(* Logix 5000 project; controller CIP_14485201 vendor 1 type 14 code 216 rev 38.11; software revision 38.01; part 10 of 12 *)
(* tags used below, declared in another part *)
   Bit : BOOL[128];   // BIT
   Integer : DINT[150];   // INTEGER
   MOA_OFF : DINT[20];   // PANELVIEW MOA OFF
   MOA_ON : DINT[20];   // PANELVIEW MOA ON
   MOA_One_Shot : BOOL[32];   // PANELVIEW MOA ONE SHOT
   MOA_Screen1_Auto : BOOL;   // PV MOA SCREEN #1 AUTO PB
   MOA_Screen1_Man_Off : BOOL;   // PV MOA SCREEN #1 OFF PB
   MOA_Screen1_Man_On : BOOL;   // PV MOA SCREEN #1 MANUAL PB
   MOA_Screen2_Auto : BOOL;   // PV MOA SCREEN #2 AUTO PB
   MOA_Screen2_Man_Off : BOOL;   // PV MOA SCREEN #2 OFF PB
   MOA_Screen2_Man_On : BOOL;   // PV MOA SCREEN #2 MANUAL PB
   MOA_Select : DINT[10];   // MAN/OFF/AUTO SELECT
   MOA_Status : DINT[10];   // MAN/OFF/AUTO STATUS
   One_Shot : BOOL[128];   // ONE SHOT ARRAY
   OpCode_Pin : DINT[5];   // OPCODE PIN ARRAY
   Panelview : INT[40];   // PANELVIEW CONTROL
   Recipe : RECIPE[41];   // RECIPES
   SCLD_Return_Temp : SCALE;   // RETURN TEMPERATURE 0-100°C
   SCLD_Rinse_Cond : SCALE;   // RINSE CONDUCTIVITY 0-10 uS/cm
   SCLD_Supply_Temp : SCALE;   // SUPPLY TEMPERATURE 0-100°C
   SCLD_Wash_Cond : SCALE;   // WASH CONDUCTIVITY 0-100 mS/cm
   SP_Return_Temp : REAL;   // CURRENT RETURN TEMP SETPOINT
   SP_Rinse_Cond : REAL;   // CURRENT RINSE CONDUCTIVITY SETPOINT
   SP_Supply_Temp : REAL;   // CURRENT SUPPLY TEMP SETPOINT
   SP_Wash_Cond : REAL;   // CURRENT WASH CONDUCTIVITY SETPOINT
   SP_Wash_Cond_Hold : REAL;   // CURRENT WASH CONDUCTIVITY SETPOINT LOW HOLD
   Subsequent_OpCode_Pin : DINT[5];   // OPCODE PIN ARRAY
   Timer : TIMER[99];   // TIMER
   Timer_Chem1_Pump : TIMER[7];   // CHEM #1 CONTROL TIMERS
   Timer_Chem2_Pump : TIMER[7];   // CHEM #2 CONTROL TIMERS
(* MainProgram, continued *)

ROUTINE _30_MAN_OFF_AUTO   (* ladder *)
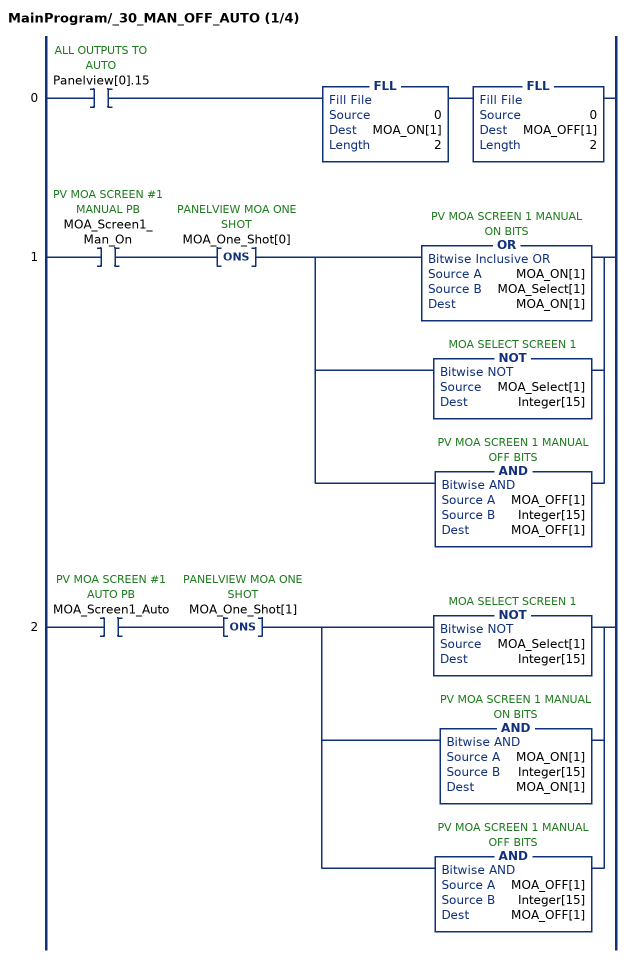
   0: XIC(Panelview[0].15)FLL(0,MOA_ON[1],2)FLL(0,MOA_OFF[1],2);
   1: XIC(MOA_Screen1_Man_On)ONS(MOA_One_Shot[0])[OR(MOA_ON[1],MOA_Select[1],MOA_ON[1]) ,NOT(MOA_Select[1],Integer[15]) ,AND(MOA_OFF[1],Integer[15],MOA_OFF[1]) ];
   2: XIC(MOA_Screen1_Auto)ONS(MOA_One_Shot[1])[NOT(MOA_Select[1],Integer[15]) ,AND(MOA_ON[1],Integer[15],MOA_ON[1]) ,AND(MOA_OFF[1],Integer[15],MOA_OFF[1]) ];
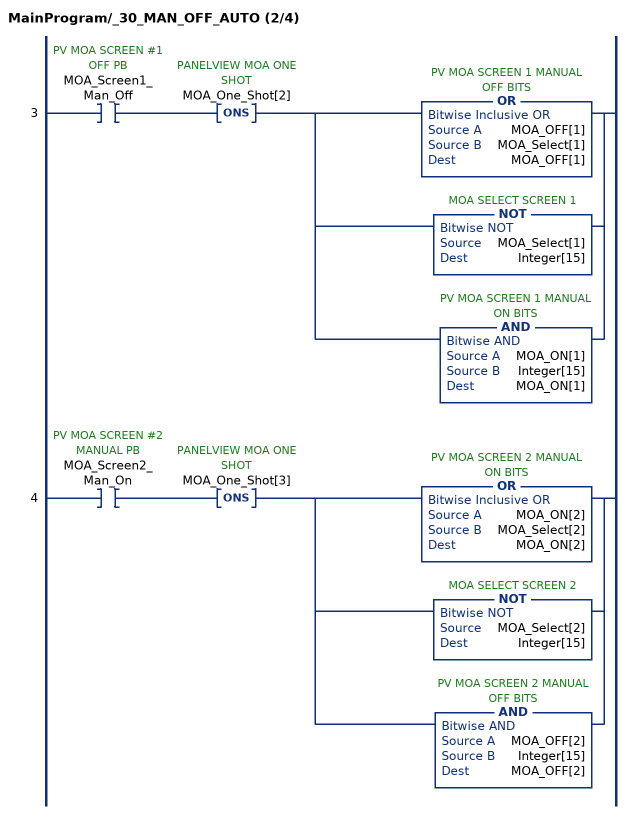
   3: XIC(MOA_Screen1_Man_Off)ONS(MOA_One_Shot[2])[OR(MOA_OFF[1],MOA_Select[1],MOA_OFF[1]) ,NOT(MOA_Select[1],Integer[15]) ,AND(MOA_ON[1],Integer[15],MOA_ON[1]) ];
   4: XIC(MOA_Screen2_Man_On)ONS(MOA_One_Shot[3])[OR(MOA_ON[2],MOA_Select[2],MOA_ON[2]) ,NOT(MOA_Select[2],Integer[15]) ,AND(MOA_OFF[2],Integer[15],MOA_OFF[2]) ];
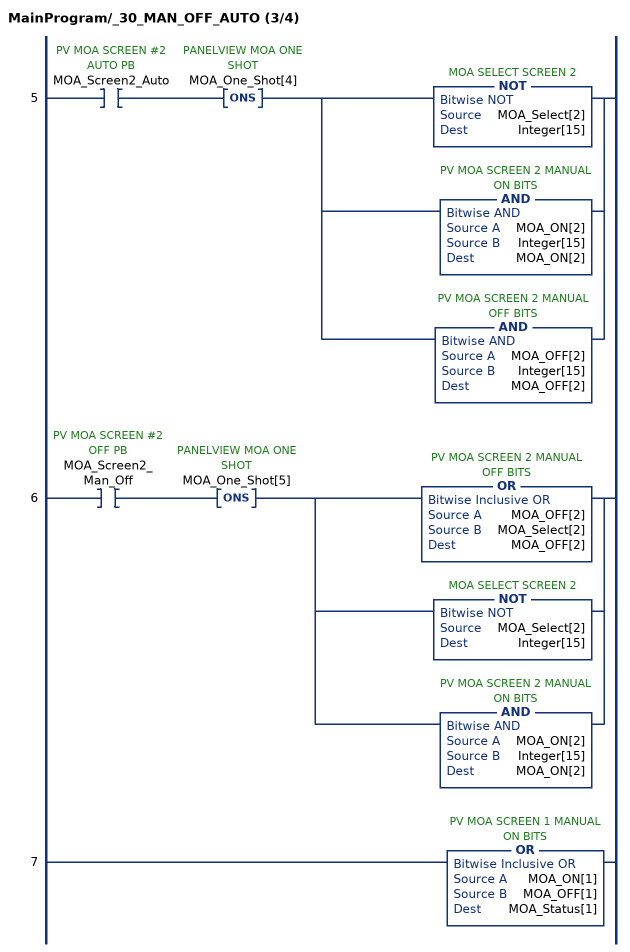
   5: XIC(MOA_Screen2_Auto)ONS(MOA_One_Shot[4])[NOT(MOA_Select[2],Integer[15]) ,AND(MOA_ON[2],Integer[15],MOA_ON[2]) ,AND(MOA_OFF[2],Integer[15],MOA_OFF[2]) ];
   6: XIC(MOA_Screen2_Man_Off)ONS(MOA_One_Shot[5])[OR(MOA_OFF[2],MOA_Select[2],MOA_OFF[2]) ,NOT(MOA_Select[2],Integer[15]) ,AND(MOA_ON[2],Integer[15],MOA_ON[2]) ];
   7: OR(MOA_ON[1],MOA_OFF[1],MOA_Status[1]);
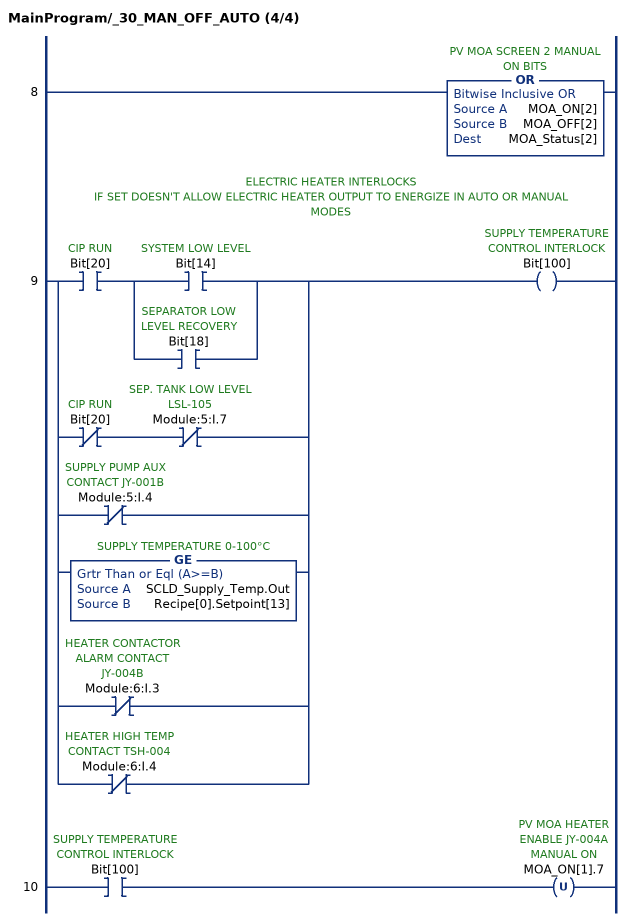
   8: OR(MOA_ON[2],MOA_OFF[2],MOA_Status[2]);
   // ELECTRIC HEATER INTERLOCKS
   // IF SET DOESN'T ALLOW ELECTRIC HEATER OUTPUT TO ENERGIZE IN AUTO OR MANUAL MODES
   9: [XIC(Bit[20]) [XIC(Bit[14]) ,XIC(Bit[18]) ] ,XIO(Bit[20]) XIO(Module:5:I.7) ,XIO(Module:5:I.4) ,GE(SCLD_Supply_Temp.Out,Recipe[0].Setpoint[13]) ,XIO(Module:6:I.3) ,XIO(Module:6:I.4) ]OTE(Bit[100]);
   10: XIC(Bit[100])OTU(MOA_ON[1].7);
END_ROUTINE

ROUTINE _86_TEMPERATURE   (* ladder *)
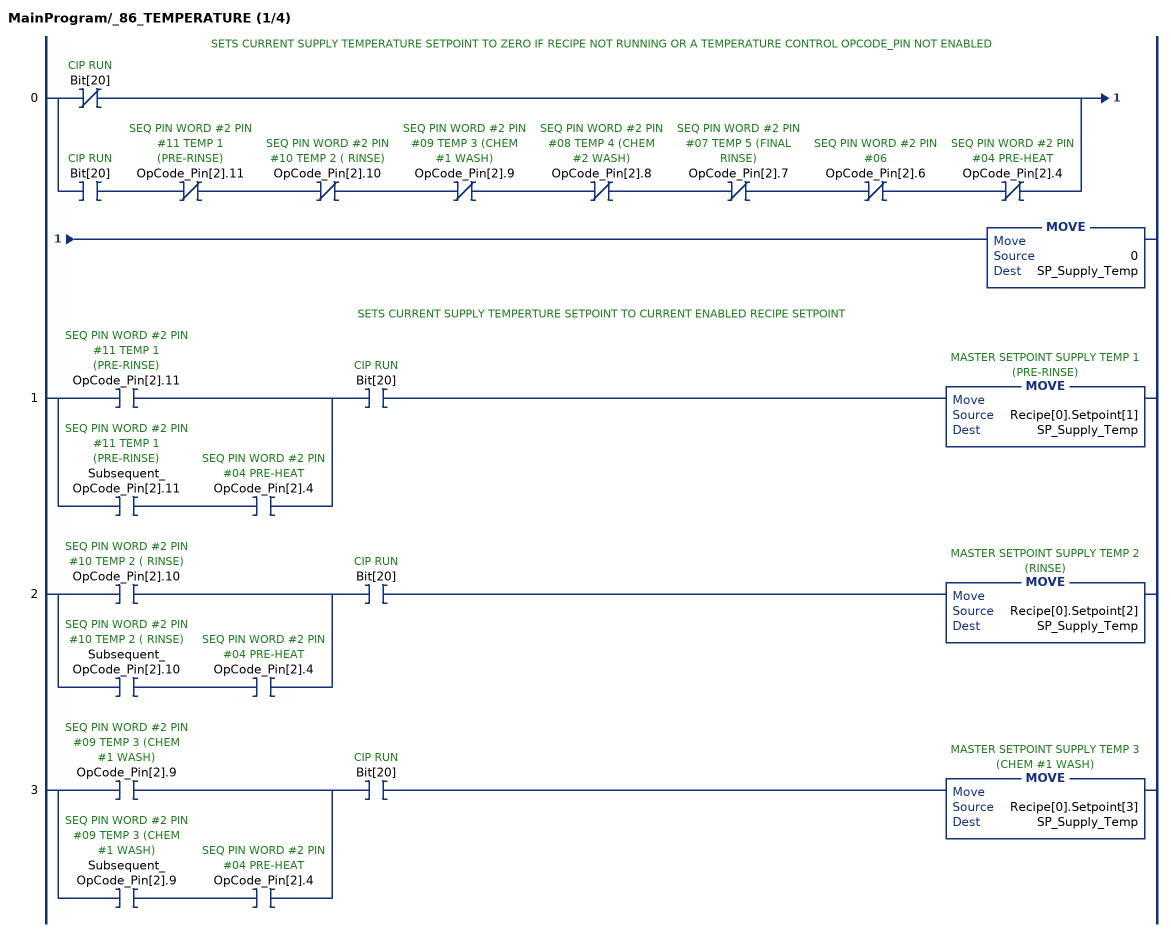
   // SETS CURRENT SUPPLY TEMPERATURE SETPOINT TO ZERO IF RECIPE NOT RUNNING OR A TEMPERATURE CONTROL OPCODE_PIN NOT ENABLED
   0: [XIO(Bit[20]) ,XIC(Bit[20]) XIO(OpCode_Pin[2].11) XIO(OpCode_Pin[2].10) XIO(OpCode_Pin[2].9) XIO(OpCode_Pin[2].8) XIO(OpCode_Pin[2].7) XIO(OpCode_Pin[2].6) XIO(OpCode_Pin[2].4) ]MOVE(0,SP_Supply_Temp);
   // SETS CURRENT SUPPLY TEMPERTURE SETPOINT TO CURRENT ENABLED RECIPE SETPOINT
   1: [XIC(OpCode_Pin[2].11) ,XIC(Subsequent_OpCode_Pin[2].11) XIC(OpCode_Pin[2].4) ]XIC(Bit[20])MOVE(Recipe[0].Setpoint[1],SP_Supply_Temp);
   2: [XIC(OpCode_Pin[2].10) ,XIC(Subsequent_OpCode_Pin[2].10) XIC(OpCode_Pin[2].4) ]XIC(Bit[20])MOVE(Recipe[0].Setpoint[2],SP_Supply_Temp);
   3: [XIC(OpCode_Pin[2].9) ,XIC(Subsequent_OpCode_Pin[2].9) XIC(OpCode_Pin[2].4) ]XIC(Bit[20])MOVE(Recipe[0].Setpoint[3],SP_Supply_Temp);
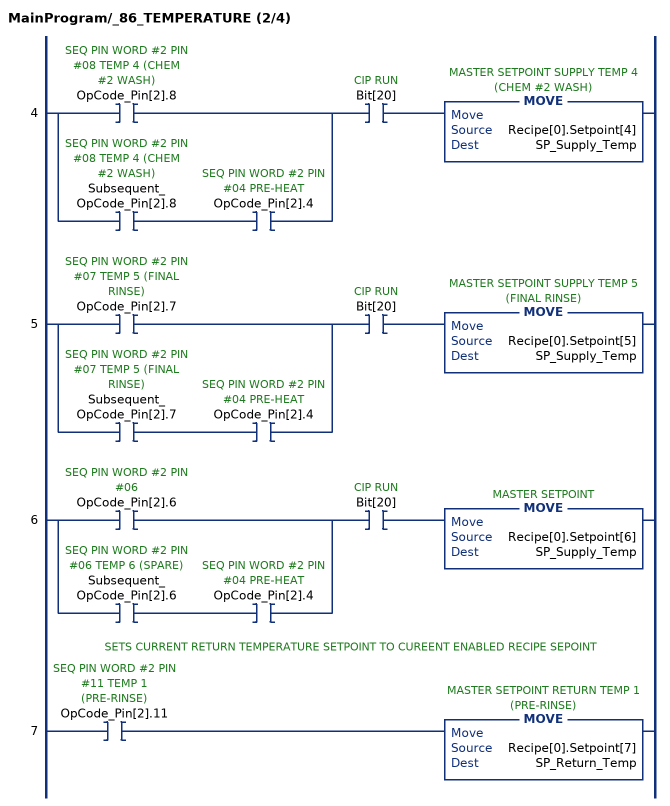
   4: [XIC(OpCode_Pin[2].8) ,XIC(Subsequent_OpCode_Pin[2].8) XIC(OpCode_Pin[2].4) ]XIC(Bit[20])MOVE(Recipe[0].Setpoint[4],SP_Supply_Temp);
   5: [XIC(OpCode_Pin[2].7) ,XIC(Subsequent_OpCode_Pin[2].7) XIC(OpCode_Pin[2].4) ]XIC(Bit[20])MOVE(Recipe[0].Setpoint[5],SP_Supply_Temp);
   6: [XIC(OpCode_Pin[2].6) ,XIC(Subsequent_OpCode_Pin[2].6) XIC(OpCode_Pin[2].4) ]XIC(Bit[20])MOVE(Recipe[0].Setpoint[6],SP_Supply_Temp);
   // SETS CURRENT RETURN TEMPERATURE SETPOINT TO CUREENT ENABLED RECIPE SEPOINT
   7: XIC(OpCode_Pin[2].11)MOVE(Recipe[0].Setpoint[7],SP_Return_Temp);
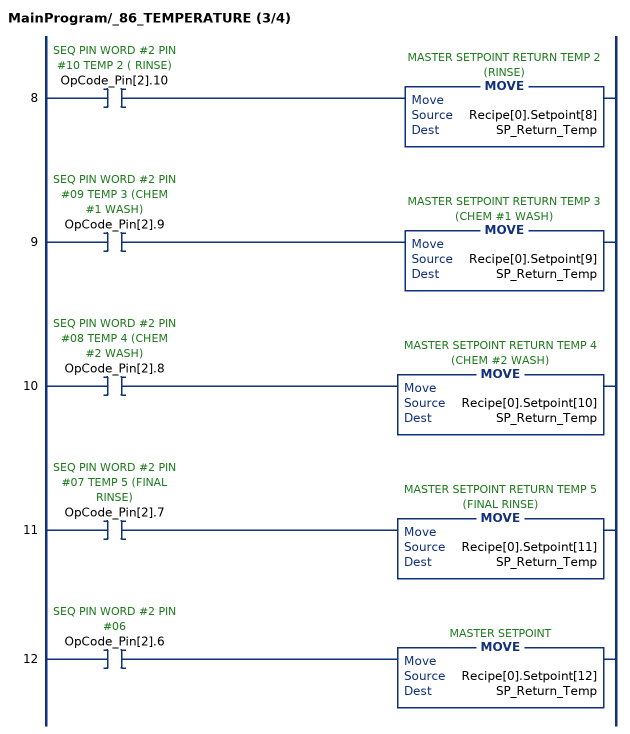
   8: XIC(OpCode_Pin[2].10)MOVE(Recipe[0].Setpoint[8],SP_Return_Temp);
   9: XIC(OpCode_Pin[2].9)MOVE(Recipe[0].Setpoint[9],SP_Return_Temp);
   10: XIC(OpCode_Pin[2].8)MOVE(Recipe[0].Setpoint[10],SP_Return_Temp);
   11: XIC(OpCode_Pin[2].7)MOVE(Recipe[0].Setpoint[11],SP_Return_Temp);
   12: XIC(OpCode_Pin[2].6)MOVE(Recipe[0].Setpoint[12],SP_Return_Temp);
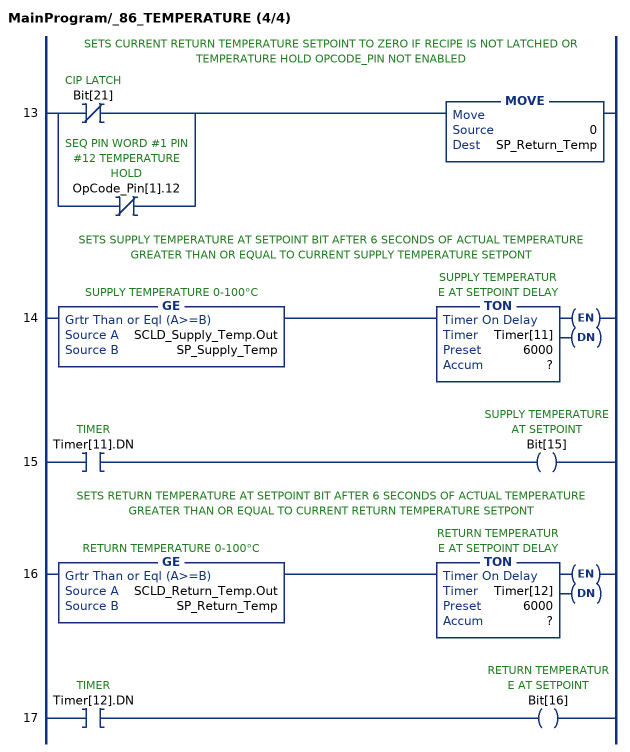
   // SETS CURRENT RETURN TEMPERATURE SETPOINT TO ZERO IF RECIPE IS NOT LATCHED OR TEMPERATURE HOLD OPCODE_PIN NOT ENABLED
   13: [XIO(Bit[21]) ,XIO(OpCode_Pin[1].12) ]MOVE(0,SP_Return_Temp);
   // SETS SUPPLY TEMPERATURE AT SETPOINT BIT AFTER 6 SECONDS OF ACTUAL TEMPERATURE GREATER THAN OR EQUAL TO CURRENT SUPPLY TEMPERATURE SETPONT
   14: GE(SCLD_Supply_Temp.Out,SP_Supply_Temp)TON(Timer[11],?,?);
   15: XIC(Timer[11].DN)OTE(Bit[15]);
   // SETS RETURN TEMPERATURE AT SETPOINT BIT AFTER 6 SECONDS OF ACTUAL TEMPERATURE GREATER THAN OR EQUAL TO CURRENT RETURN TEMPERATURE SETPONT
   16: GE(SCLD_Return_Temp.Out,SP_Return_Temp)TON(Timer[12],?,?);
   17: XIC(Timer[12].DN)OTE(Bit[16]);
END_ROUTINE

ROUTINE _87_CHEM1_PUMP   (* ladder *)
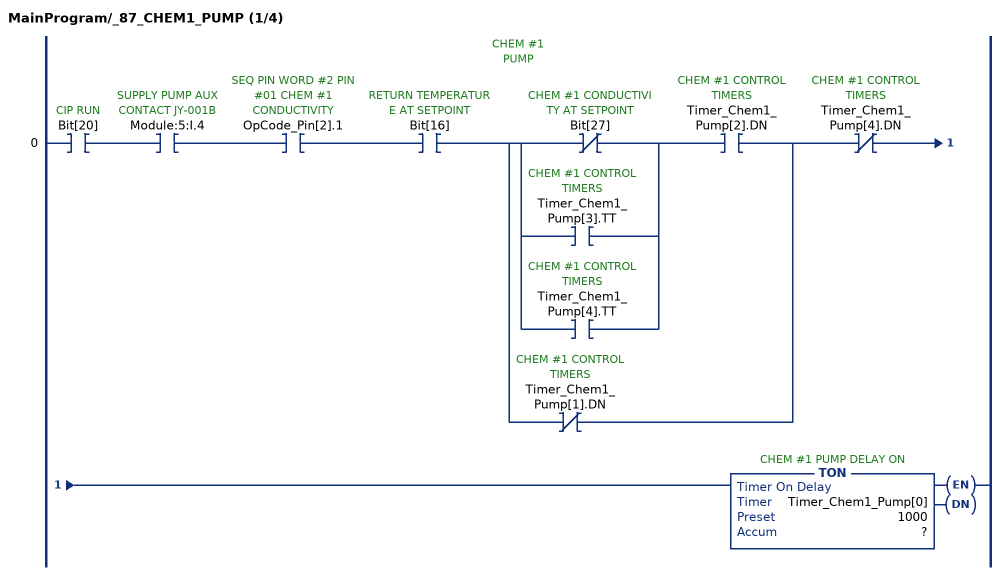
   // CHEM #1
   // PUMP
   0: XIC(Bit[20])XIC(Module:5:I.4)XIC(OpCode_Pin[2].1)XIC(Bit[16])[[XIO(Bit[27]) ,XIC(Timer_Chem1_Pump[3].TT) ,XIC(Timer_Chem1_Pump[4].TT) ] XIC(Timer_Chem1_Pump[2].DN) ,XIO(Timer_Chem1_Pump[1].DN) ]XIO(Timer_Chem1_Pump[4].DN)TON(Timer_Chem1_Pump[0],?,?);
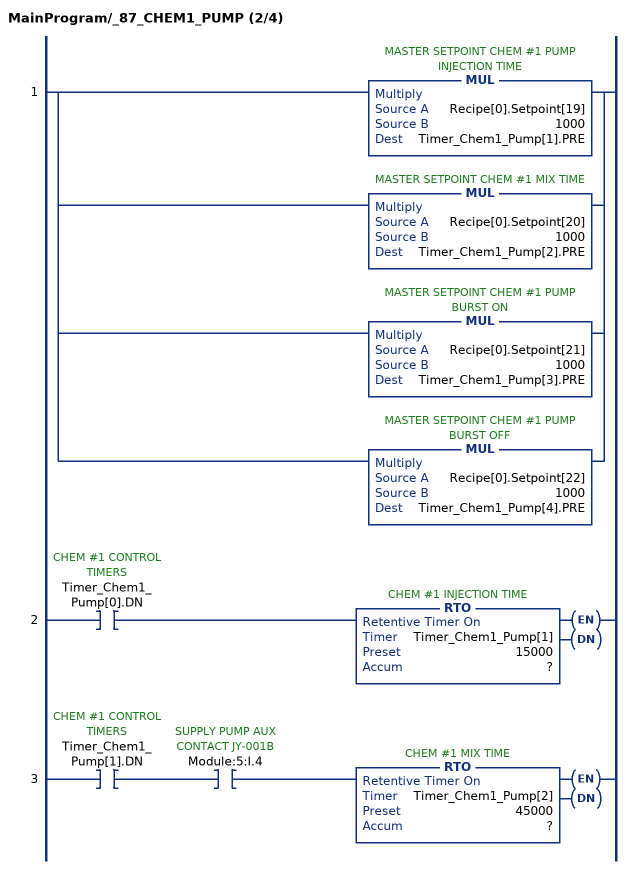
   1: [MUL(Recipe[0].Setpoint[19],1000,Timer_Chem1_Pump[1].PRE) ,MUL(Recipe[0].Setpoint[20],1000,Timer_Chem1_Pump[2].PRE) ,MUL(Recipe[0].Setpoint[21],1000,Timer_Chem1_Pump[3].PRE) ,MUL(Recipe[0].Setpoint[22],1000,Timer_Chem1_Pump[4].PRE) ];
   2: XIC(Timer_Chem1_Pump[0].DN)RTO(Timer_Chem1_Pump[1],?,?);
   3: XIC(Timer_Chem1_Pump[1].DN)XIC(Module:5:I.4)RTO(Timer_Chem1_Pump[2],?,?);
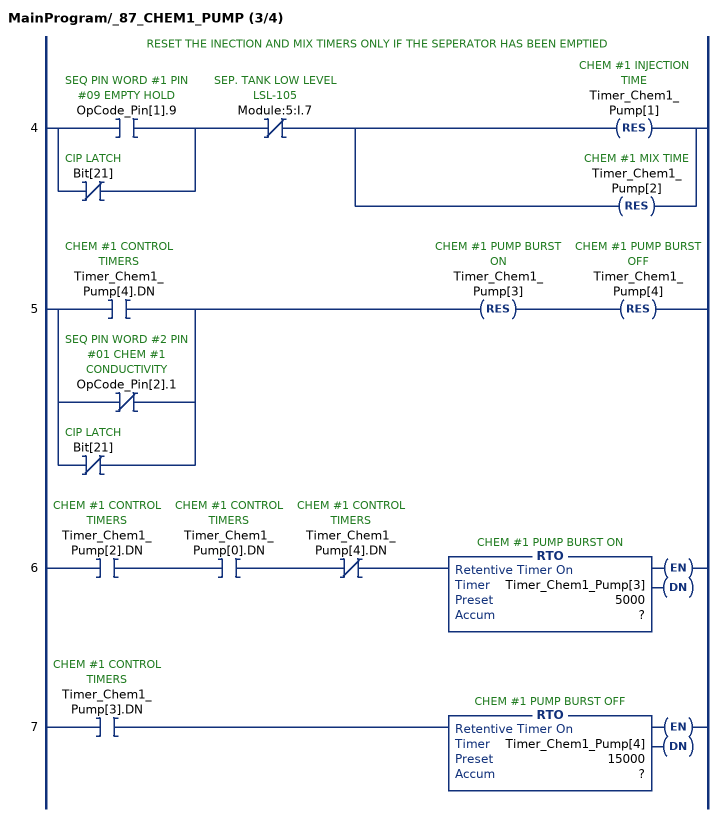
   // RESET THE INECTION AND MIX TIMERS ONLY IF THE SEPERATOR HAS BEEN EMPTIED
   4: [XIC(OpCode_Pin[1].9) ,XIO(Bit[21]) ]XIO(Module:5:I.7)[RES(Timer_Chem1_Pump[1]) ,RES(Timer_Chem1_Pump[2]) ];
   5: [XIC(Timer_Chem1_Pump[4].DN) ,XIO(OpCode_Pin[2].1) ,XIO(Bit[21]) ]RES(Timer_Chem1_Pump[3])RES(Timer_Chem1_Pump[4]);
   6: XIC(Timer_Chem1_Pump[2].DN)XIC(Timer_Chem1_Pump[0].DN)XIO(Timer_Chem1_Pump[4].DN)RTO(Timer_Chem1_Pump[3],?,?);
   7: XIC(Timer_Chem1_Pump[3].DN)RTO(Timer_Chem1_Pump[4],?,?);
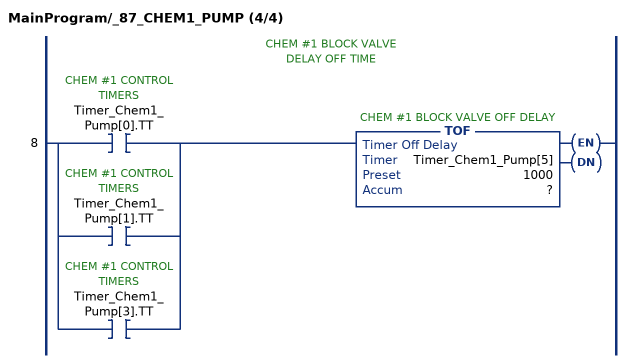
   // CHEM #1 BLOCK VALVE
   //  DELAY OFF TIME
   8: [XIC(Timer_Chem1_Pump[0].TT) ,XIC(Timer_Chem1_Pump[1].TT) ,XIC(Timer_Chem1_Pump[3].TT) ]TOF(Timer_Chem1_Pump[5],?,?);
END_ROUTINE

ROUTINE _87_CHEM2_PUMP   (* ladder *)
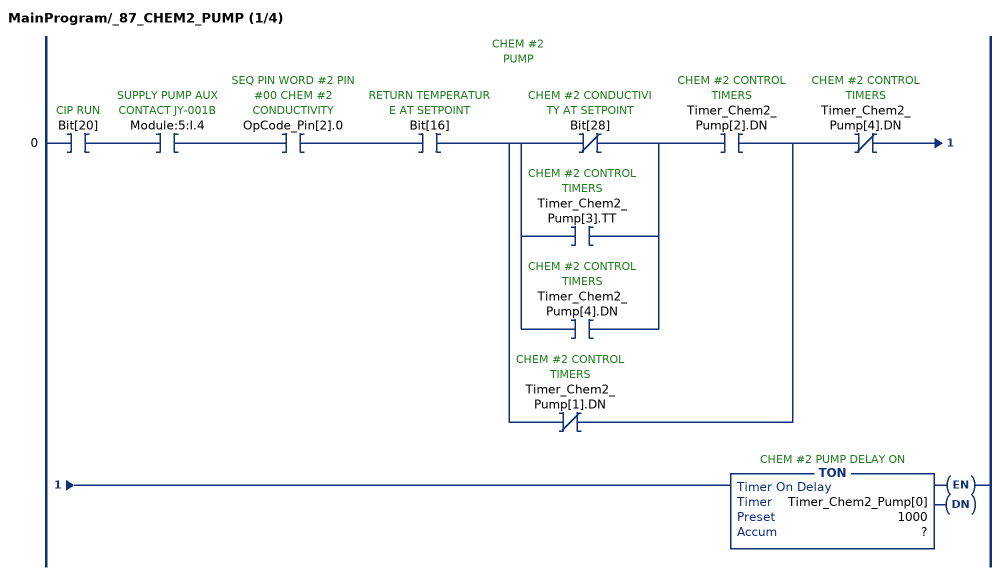
   // CHEM #2
   // PUMP
   0: XIC(Bit[20])XIC(Module:5:I.4)XIC(OpCode_Pin[2].0)XIC(Bit[16])[[XIO(Bit[28]) ,XIC(Timer_Chem2_Pump[3].TT) ,XIC(Timer_Chem2_Pump[4].DN) ] XIC(Timer_Chem2_Pump[2].DN) ,XIO(Timer_Chem2_Pump[1].DN) ]XIO(Timer_Chem2_Pump[4].DN)TON(Timer_Chem2_Pump[0],?,?);
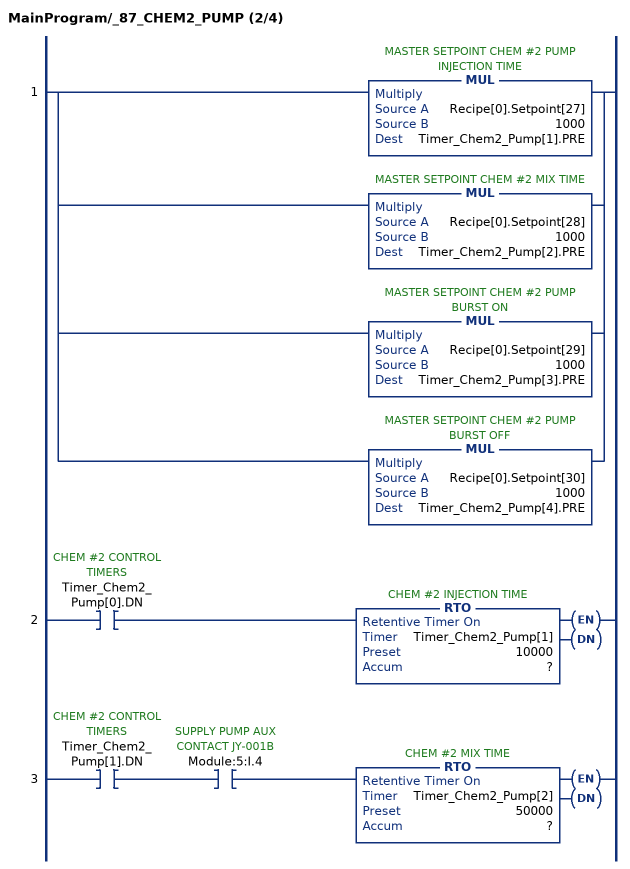
   1: [MUL(Recipe[0].Setpoint[27],1000,Timer_Chem2_Pump[1].PRE) ,MUL(Recipe[0].Setpoint[28],1000,Timer_Chem2_Pump[2].PRE) ,MUL(Recipe[0].Setpoint[29],1000,Timer_Chem2_Pump[3].PRE) ,MUL(Recipe[0].Setpoint[30],1000,Timer_Chem2_Pump[4].PRE) ];
   2: XIC(Timer_Chem2_Pump[0].DN)RTO(Timer_Chem2_Pump[1],?,?);
   3: XIC(Timer_Chem2_Pump[1].DN)XIC(Module:5:I.4)RTO(Timer_Chem2_Pump[2],?,?);
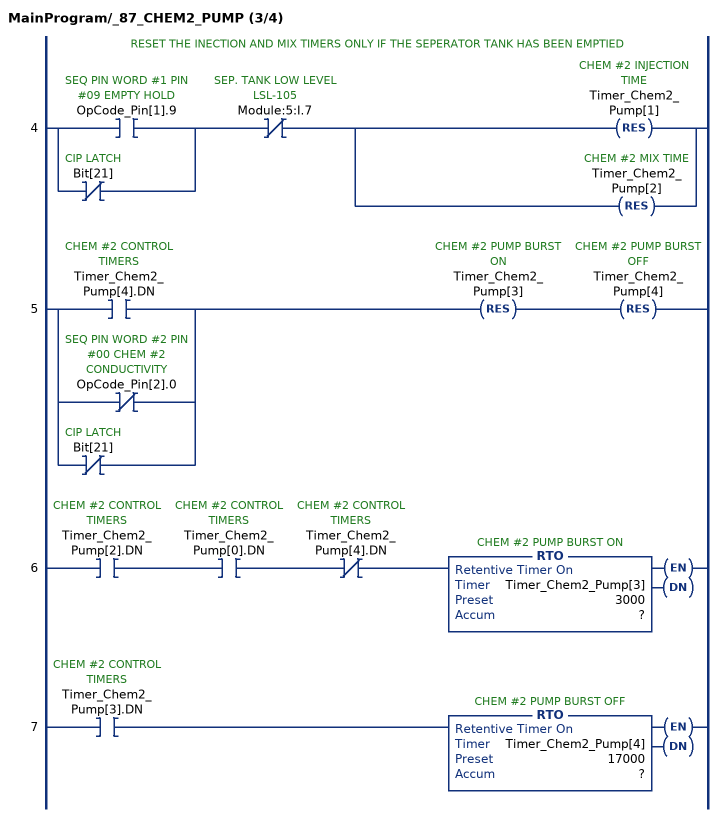
   // RESET THE INECTION AND MIX TIMERS ONLY IF THE SEPERATOR TANK HAS BEEN EMPTIED
   4: [XIC(OpCode_Pin[1].9) ,XIO(Bit[21]) ]XIO(Module:5:I.7)[RES(Timer_Chem2_Pump[1]) ,RES(Timer_Chem2_Pump[2]) ];
   5: [XIC(Timer_Chem2_Pump[4].DN) ,XIO(OpCode_Pin[2].0) ,XIO(Bit[21]) ]RES(Timer_Chem2_Pump[3])RES(Timer_Chem2_Pump[4]);
   6: XIC(Timer_Chem2_Pump[2].DN)XIC(Timer_Chem2_Pump[0].DN)XIO(Timer_Chem2_Pump[4].DN)RTO(Timer_Chem2_Pump[3],?,?);
   7: XIC(Timer_Chem2_Pump[3].DN)RTO(Timer_Chem2_Pump[4],?,?);
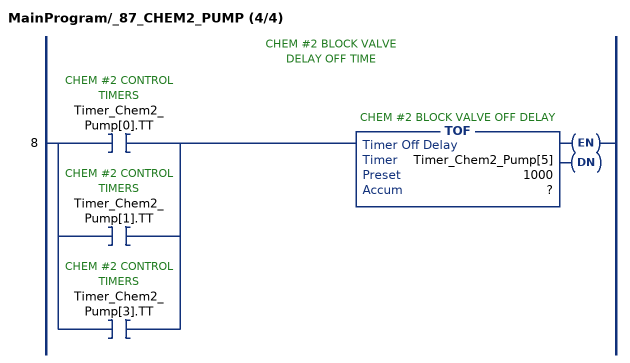
   // CHEM #2 BLOCK VALVE
   //  DELAY OFF TIME
   8: [XIC(Timer_Chem2_Pump[0].TT) ,XIC(Timer_Chem2_Pump[1].TT) ,XIC(Timer_Chem2_Pump[3].TT) ]TOF(Timer_Chem2_Pump[5],?,?);
END_ROUTINE

ROUTINE _87_CONDUCTIVITY   (* ladder *)
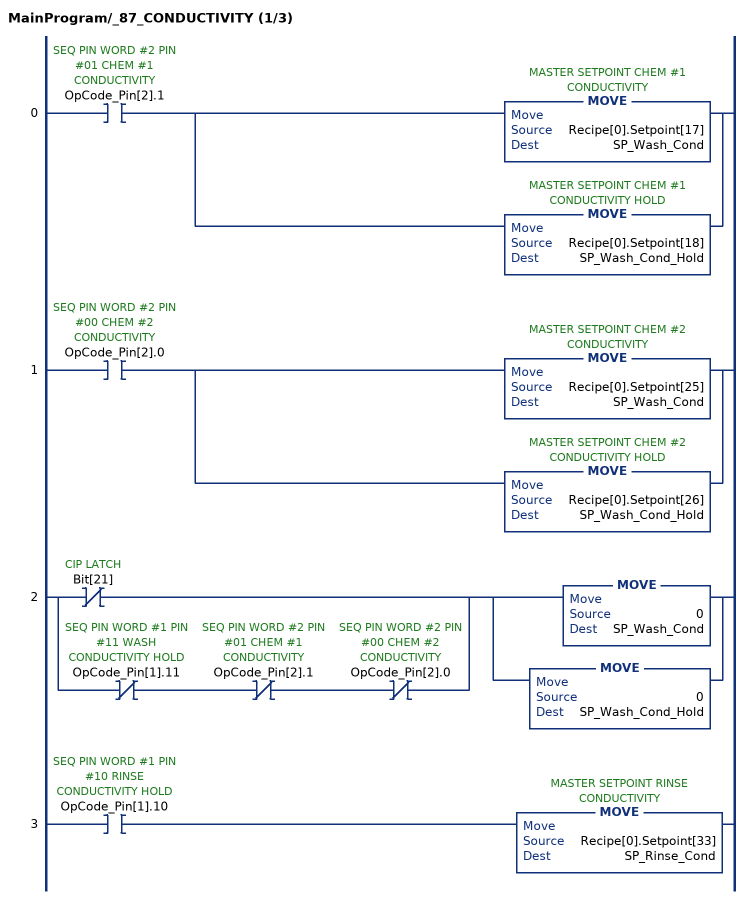
   0: XIC(OpCode_Pin[2].1)[MOVE(Recipe[0].Setpoint[17],SP_Wash_Cond) ,MOVE(Recipe[0].Setpoint[18],SP_Wash_Cond_Hold) ];
   1: XIC(OpCode_Pin[2].0)[MOVE(Recipe[0].Setpoint[25],SP_Wash_Cond) ,MOVE(Recipe[0].Setpoint[26],SP_Wash_Cond_Hold) ];
   2: [XIO(Bit[21]) ,XIO(OpCode_Pin[1].11) XIO(OpCode_Pin[2].1) XIO(OpCode_Pin[2].0) ][MOVE(0,SP_Wash_Cond) ,MOVE(0,SP_Wash_Cond_Hold) ];
   3: XIC(OpCode_Pin[1].10)MOVE(Recipe[0].Setpoint[33],SP_Rinse_Cond);
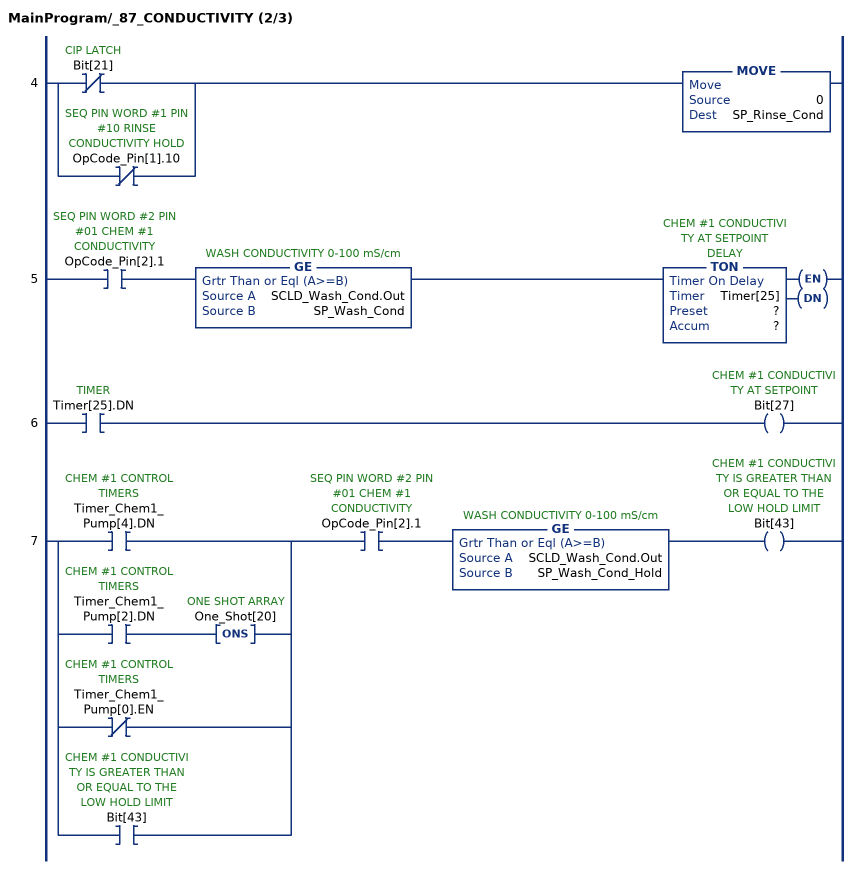
   4: [XIO(Bit[21]) ,XIO(OpCode_Pin[1].10) ]MOVE(0,SP_Rinse_Cond);
   5: XIC(OpCode_Pin[2].1)GE(SCLD_Wash_Cond.Out,SP_Wash_Cond)TON(Timer[25],?,?);
   6: XIC(Timer[25].DN)OTE(Bit[27]);
   7: [XIC(Timer_Chem1_Pump[4].DN) ,XIC(Timer_Chem1_Pump[2].DN) ONS(One_Shot[20]) ,XIO(Timer_Chem1_Pump[0].EN) ,XIC(Bit[43]) ]XIC(OpCode_Pin[2].1)GE(SCLD_Wash_Cond.Out,SP_Wash_Cond_Hold)OTE(Bit[43]);
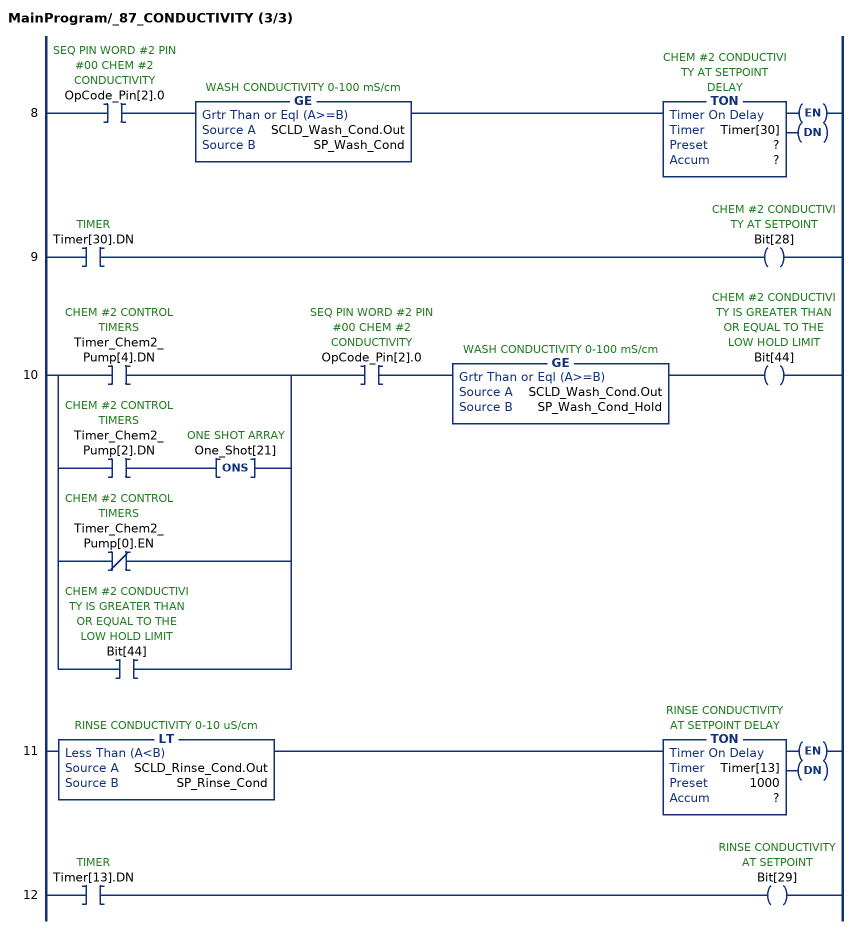
   8: XIC(OpCode_Pin[2].0)GE(SCLD_Wash_Cond.Out,SP_Wash_Cond)TON(Timer[30],?,?);
   9: XIC(Timer[30].DN)OTE(Bit[28]);
   10: [XIC(Timer_Chem2_Pump[4].DN) ,XIC(Timer_Chem2_Pump[2].DN) ONS(One_Shot[21]) ,XIO(Timer_Chem2_Pump[0].EN) ,XIC(Bit[44]) ]XIC(OpCode_Pin[2].0)GE(SCLD_Wash_Cond.Out,SP_Wash_Cond_Hold)OTE(Bit[44]);
   11: LT(SCLD_Rinse_Cond.Out,SP_Rinse_Cond)TON(Timer[13],?,?);
   12: XIC(Timer[13].DN)OTE(Bit[29]);
END_ROUTINE
